Fanuc KAREL source: kd00026.KL

-- PROVISIONAL review KL for V1013-1; original PC SHA256 f1143c8eba3c43c5e00a86c35554b752bd82744ce8965ab50226d67fe0a748a7
-- Incomplete behavior may be omitted. Consult companion uncertainty JSON. Do not deploy.
PROGRAM KD00026
%NOLOCKGROUP
VAR
  I : INTEGER
  J : INTEGER
  B : BOOLEAN
  R : REAL
  S : STRING[80]
BEGIN
  -- UNRESOLVED_PC offsets 5-24; opcodes 9D,81,18,9D,1B,9D,12,22,9D,13,04
  -- UNRESOLVED_PC offsets 29-33; opcodes 7F
END KD00026
